Fanuc KAREL source: kb00015.KL

-- PROVISIONAL review KL for V1013-1; original PC SHA256 b825d03005622cd6e51f5b60d47270ff36f462a81b51c471a1ce00aec02e9054
-- Incomplete behavior may be omitted. Consult companion uncertainty JSON. Do not deploy.
PROGRAM KB00015
%NOLOCKGROUP
BEGIN
  -- UNRESOLVED_PC offsets 5-14; opcodes 3F,75
  -- UNRESOLVED_PC offsets 19-26; opcodes 9D,23
  -- UNRESOLVED_PC offsets 31-49; opcodes 27,22,2A,22,31
  -- UNRESOLVED_PC offsets 54-58; opcodes 7F
END KB00015
